(* IEC 61131-3 sources: plcassist-cli/packages/volt-lsp-iec/test-corpus/bakon-nano/Device/Plc Logic/Application/Library Manager/L_TF2P_TechModulesFollowingPositioning, 28 files *)

(* ---- L_TF2P_CONSTANTS.gvl ---- *)
VAR_GLOBAL
	GC_DWCHECKIDTAPPETREF : DWORD := 16#DC34;
	GC_LREPSILON : LREAL := 1E-06;
	GC_POSITIVE_LIMIT_32BIT : LREAL := 2147483647;
	GC_NEGATIVE_LIMIT_32BIT : LREAL := -2147483647;
	GC_PI : LREAL := 3.1415926535897931;
END_VAR

(* ---- L_TF2P_IACCESSPOINTS.itf ---- *)
INTERFACE L_TF2P_IACCESSPOINTS
END_INTERFACE

METHOD GET_PAP : POINTER TO L_TF2P_scAP_TM_TablePositioningBase
END_METHOD

(* ---- L_TF2P_ICONNECTORTABLEPOS.itf ---- *)
INTERFACE L_TF2P_ICONNECTORTABLEPOS
END_INTERFACE

(* ---- L_TF2P_ITABLEPOSITIONINGBASE.itf ---- *)
INTERFACE L_TF2P_ITABLEPOSITIONINGBASE
END_INTERFACE

METHOD PROFILEGENERATOR
VAR_INPUT
	ITFTECHMODULE : L_TF2P_ITablePositioningBase;
	XEXECUTE : BOOL;
	XCONTINUOUSUPDATE : BOOL;
	LRPOSITION : LREAL;
	LRVELOCITY : LREAL;
	LRENDVELOCITY : LREAL;
	LRACCELERATION : LREAL;
	LRDECELERATION : LREAL;
	LRJERK : LREAL;
	XPOSMODE : BOOL;
	EDIRECTION : MC_DIRECTION;
	EFUNCTIONTYP : L_MC1P_TypeFunction;
END_VAR
VAR_OUTPUT
	XDONE : BOOL;
	XBUSY : BOOL;
	XACTIVE : BOOL;
	XCOMMANDABORTED : BOOL;
	XERROR : BOOL;
	EERRORID : L_IE1P_Error;
END_VAR
VAR_IN_OUT
	AXIS : AXIS_REF;
END_VAR
END_METHOD

(* ---- GETBOOLEANPROPERTY.fun ---- *)
FUNCTION GETBOOLEANPROPERTY : BOOL
VAR_INPUT
	STKEY : WSTRING;
END_VAR
END_FUNCTION

(* ---- GETCOMPANY.fun ---- *)
FUNCTION GETCOMPANY : WSTRING
END_FUNCTION

(* ---- GETNUMBERPROPERTY.fun ---- *)
FUNCTION GETNUMBERPROPERTY : DINT
VAR_INPUT
	STKEY : WSTRING;
END_VAR
END_FUNCTION

(* ---- GETTEXTPROPERTY.fun ---- *)
FUNCTION GETTEXTPROPERTY : WSTRING
VAR_INPUT
	STKEY : WSTRING;
END_VAR
END_FUNCTION

(* ---- GETTEXTPROPERTY2.fun ---- *)
FUNCTION GETTEXTPROPERTY2 : POINTER TO WSTRING
VAR_INPUT
	STKEY : WSTRING;
END_VAR
END_FUNCTION

(* ---- GETTITLE.fun ---- *)
FUNCTION GETTITLE : WSTRING
END_FUNCTION

(* ---- GETVERSION.fun ---- *)
FUNCTION GETVERSION : VERSION
END_FUNCTION

(* ---- GETVERSIONPROPERTY.fun ---- *)
FUNCTION GETVERSIONPROPERTY : VERSION
VAR_INPUT
	STKEY : WSTRING;
END_VAR
END_FUNCTION

(* ---- L_TF2P_CHECKEXTERNALBYLIMITER.fun ---- *)
FUNCTION L_TF2P_CHECKEXTERNALBYLIMITER : BOOL
VAR_INPUT
	DWLIMITERCONTROL : DWORD;
END_VAR
VAR_IN_OUT
	AXIS : AXIS_REF;
END_VAR
END_FUNCTION

(* ---- L_TF2P_GETSTARTMOVETOTARGETPOS.fun ---- *)
FUNCTION L_TF2P_GETSTARTMOVETOTARGETPOS : BOOL
VAR_INPUT
	MASTERVALUES : L_MC1P_IAXIS_REF_MASTERVALUES;
	LRSYNCDEC : LREAL;
	LRSYNCJERK : LREAL;
	LRTARGETPOS : LREAL;
END_VAR
VAR_IN_OUT
	AXIS : AXIS_REF;
END_VAR
END_FUNCTION

(* ---- L_TF2P_POSITIONINSIDEWINDOW.fun ---- *)
FUNCTION L_TF2P_POSITIONINSIDEWINDOW : BOOL
VAR_INPUT
	LRPOSIN : LREAL;
	LRLOWERWINDOW : LREAL;
	LRUPPERWINDOW : LREAL;
END_VAR
VAR_OUTPUT
	XERROR : BOOL := FALSE;
END_VAR
VAR_IN_OUT
	AXIS : AXIS_REF;
END_VAR
END_FUNCTION

(* ---- GLOBALTEXTLIST.fb ---- *)
FUNCTION_BLOCK GLOBALTEXTLIST
VAR
	M_TEXTLISTFILE : STRING(255);
	_STNAMESPACE : STRING;
END_VAR
END_FUNCTION_BLOCK

(* ---- L_TB2A_PROFILEMANAGER.fb ---- *)
FUNCTION_BLOCK L_TB2A_PROFILEMANAGER
VAR_INPUT
	XEXECUTE : BOOL;
	XABORT : BOOL;
	WSTARTNUMBER : WORD;
	XNEXTPROFILE : BOOL;
END_VAR
VAR_OUTPUT
	XBUSY : BOOL;
	XDONE : BOOL;
	XABORTED : BOOL;
	XERROR : BOOL;
	EERRORID : L_IE1P_Error;
	XPROFILEERROR : BOOL;
	EPROFILEERRORID : L_IE1P_Error;
	WACTPROFILE : WORD;
	PACTPROFILE : POINTER TO L_TF2P_scPositionProfile;
	XHASNEXT : BOOL;
	XRTRIG : BOOL;
	EPROFILETYPE : L_MC1P_TypeFunction;
	XMOVEABS : BOOL;
	XMOVEREL : BOOL;
	XMOVEVEL : BOOL;
	XMOVECONTABS : BOOL;
	XMOVECONTREL : BOOL;
	XTPINSIDEWINDOW : BOOL;
	XTPOUTSIDEWINDOW : BOOL;
	XTPMISSED : BOOL;
	EDIRECTION : MC_DIRECTION;
END_VAR
VAR_IN_OUT
	ASCPROFILES : ARRAY [1..15] OF L_TF2P_scPositionProfile;
	SCTPRECDATA : L_MC1P_TpReceiveData;
	AXIS : AXIS_REF;
END_VAR
VAR
	_MODEL : L_UBUP_BehaviourModel_ETrigA;
	_XNEXTPROFILETRIG : R_TRIG;
	_XTPPROFILE : R_TRIG;
	LRTP_RELDIFF : LREAL;
	XTPWINDOWOPENED : BOOL;
	XTPWINDOWOPEN : BOOL;
	XTP_REL_PROFILEACTIVE : BOOL;
END_VAR
END_FUNCTION_BLOCK

METHOD CYCLICACTION
VAR_INPUT
	ITFTIMINGCONTROLLER : L_UBUP_ITimingController;
END_VAR
VAR_OUTPUT
	XCOMPLETE : BOOL;
	XABORT : BOOL;
	IERRORID : INT;
END_VAR
END_METHOD

METHOD FINALIZEACTION
VAR_INPUT
	XABORTPROPOSED : BOOL;
	IERRORIDPROPOSED : INT;
END_VAR
VAR_OUTPUT
	XCOMPLETE : BOOL;
	XABORT : BOOL;
	IERRORID : INT;
END_VAR
END_METHOD

METHOD RESETACTION
VAR_OUTPUT
	XCOMPLETE : BOOL;
END_VAR
END_METHOD

METHOD STARTACTION
VAR_OUTPUT
	XCOMPLETE : BOOL;
	IERRORID : INT;
END_VAR
END_METHOD

METHOD FB_INIT : BOOL
VAR_INPUT
	BINITRETAINS : BOOL;
	BINCOPYCODE : BOOL;
END_VAR
END_METHOD

METHOD GET_POSITIONINGMODE
VAR_OUTPUT
	EERRORID : L_IE1P_Error;
END_VAR
END_METHOD

METHOD GET_PROFILE
END_METHOD

METHOD GET_TPDETECTION
VAR_OUTPUT
	EERRORID : L_IE1P_Error;
END_VAR
END_METHOD

(* ---- L_TF2P_CONDITIONPROFILEMANAGER.fb ---- *)
FUNCTION_BLOCK L_TF2P_CONDITIONPROFILEMANAGER EXTENDS L_UBUP_ConditionBase
VAR_INPUT
	EPOSITIONINGMODE : L_TF2P_ePositioningMode;
	EINVALIDPROFILEID : L_IE1P_Error;
	EACTSTATE : L_TB2P_States;
END_VAR
VAR_IN_OUT
	AXIS : AXIS_REF;
END_VAR
END_FUNCTION_BLOCK

METHOD VERIFY : BOOL
VAR_OUTPUT
	XCONDITIONERROR : BOOL;
	EERRORIDPROPOSED : L_IE1P.L_IE1P_Error;
END_VAR
END_METHOD

(* ---- L_TF2P_CONTROLUNIT_ACTUALSPEED.fb ---- *)
FUNCTION_BLOCK L_TF2P_CONTROLUNIT_ACTUALSPEED
VAR_INPUT
	XENABLE : BOOL := FALSE;
	XENABLEOPERATION : BOOL := FALSE;
	XSPEEDCONTROL : BOOL := FALSE;
	SCPROFILELIMITS : L_TF2P_scProfileLimits;
	XENABLEEXTVEL : BOOL := FALSE;
	LREXTVEL : LREAL := 0;
	XENABLEEXTACCDECJERK : BOOL := FALSE;
	LREXTACC : LREAL := 0;
	LREXTDEC : LREAL := 0;
	LREXTJERK : LREAL := 0;
	XENABLEEXTTRQ : BOOL := FALSE;
	LREXTTRQ : LREAL := 0;
	XFASTSLOW : BOOL;
	XINVERTDIRECTION : BOOL;
	SCPROFILEACTUALSPEED : L_TF2P_scProfileDataState_int;
	XBRAKEISUSED : BOOL := FALSE;
	XBRAKERELEASED : BOOL := FALSE;
	ETMSTATES : L_TB2P_States;
	XAXISWARNING : BOOL;
	XTMERROR : BOOL;
	XSTO : BOOL;
	XAXISENABLED : BOOL := FALSE;
	XAXISREADY : BOOL := FALSE;
END_VAR
VAR_OUTPUT
	XENABLED : BOOL := FALSE;
	XBUSY : BOOL := FALSE;
	SCCONTROLUNIT : L_TF2P_scControlUnit;
	XERROR : BOOL;
	EERRORID : L_IE1P_Error;
	XEXTVELACTIVE : BOOL;
	XEXTTRQACTIVE : BOOL;
	XEXTACCDECJERKACTIVE : BOOL := FALSE;
	XMOVEVELEXECUTE : BOOL;
	XABORTOUT : BOOL;
	ESETDIRECTION : L_MC1P.MC_DIRECTION;
END_VAR
VAR_IN_OUT
	XNEWCOMMAND : BOOL;
END_VAR
VAR
	XNOTFIRSTCYCLE : BOOL := FALSE;
	XSPEEDCONTROL_OLD : BOOL;
END_VAR
END_FUNCTION_BLOCK

(* ---- L_TF2P_FOLLOWSETVALUESBASE.fb ---- *)
FUNCTION_BLOCK L_TF2P_FOLLOWSETVALUESBASE EXTENDS L_TB2P_TechModuleBase
VAR_INPUT
	XENABLE : BOOL;
	XENABLEOPERATION : BOOL;
	XRESETERROR : BOOL;
	XQSPAPPLICATION : BOOL;
	XABORT : BOOL;
	XJOGPOS : BOOL;
	XJOGNEG : BOOL;
	XHOMEEXECUTE : BOOL;
	LROVERRIDE : LREAL := 1;
	SCCTRLBASICMOTION : L_TB2P_scCtrlBasicMotion;
	SCPAR : L_TF2P_scPar_FollowSetValuesBase;
	SCACCESSPOINTS : L_TF2P_scAP_FollowSetValuesBase;
	XFOLLOWSETVALUES : BOOL;
	LRSETVELOCITY : LREAL;
	LRSETTORQUE : LREAL;
END_VAR
VAR_OUTPUT
	XREADYFOROPERATION : BOOL;
	XOPERATIONENABLED : BOOL;
	XREADYFORMOTION : BOOL;
	XERROR : BOOL;
	XWARNING : BOOL;
	EERRORID : L_IE1P_Error;
	XSTOACTIVE : BOOL;
	XQSPACTIVE : BOOL;
	XABORTBUSY : BOOL;
	XABORTDONE : BOOL;
	XJOGGINGBUSY : BOOL;
	XHOMINGBUSY : BOOL;
	XHOMINGDONE : BOOL;
	XISHOMED : BOOL;
	ETMSTATE : L_TB2P_States := L_TB2P_States.DISABLED;
	SCSTATUSBASICMOTION : L_TB2P_scStatusBasicMotion;
	LRACTVEL : LREAL;
	LRSETVELOUT : LREAL;
	LRACTPOS : LREAL;
	LRSETPOSOUT : LREAL;
	LRACTFOLLOWINGERROR : LREAL;
	SCSIGNALFLOW : L_TF2P_scSF_FollowSetValuesBase;
	XFOLLOWVELOCITYBUSY : BOOL;
	XFOLLOWTORQUEBUSY : BOOL;
	XVELLIMITACTIVE : BOOL;
	XACCDECLIMITACTIVE : BOOL;
	XTORQUEINTARGET : BOOL;
	LRACTTORQUE : LREAL;
	LRSETTORQUEOUT : LREAL;
END_VAR
VAR_IN_OUT
	AXIS : AXIS_REF;
END_VAR
VAR
	TM_INT : L_TF2P_TM_FollowSetValuesBase := STRUCT(ModuleHandler := ModuleHandler);
	XENABLE_OLD : BOOL;
	_UICALLMFUNIDXINPUT : UINT := 1;
	_UICALLMFUNIDXOUTPUT : UINT := 1;
	_ASCINPUT : ARRAY [1.._MCCall.c_BufferDepthInput] OF L_TF2P_FollowSetValuesBaseIn;
	_ASCOUTPUT : ARRAY [1.._MCCall.c_BufferDepthOutput] OF L_TF2P_FollowSetValuesBaseOut;
	_ASCPARCORE : ARRAY [1.._MCCall.c_BufferDepthInput] OF L_TF2P_scPar_FollowSetValuesBase;
	_ASCACCESSPOINTSCORE : ARRAY [1.._MCCall.c_BufferDepthInput] OF L_TF2P_scAP_FollowSetValuesBase;
	_ASCSIGNALFLOWCORE : ARRAY [1.._MCCall.c_BufferDepthOutput] OF L_TF2P_scSF_FollowSetValuesBase;
	_MCCALL : L_UM1P_MCCall;
	SCPAR_INT : L_TF2P_scPar_FollowSetValuesBase;
	_SCINPUTVISU : L_TF2P_FollowSetValuesBaseIn;
	_PSCINPUTVISU : POINTER TO L_TF2P_FollowSetValuesBaseIn := ADR(_scInputVisu);
	_PSCOUTPUTVISU : POINTER TO L_TF2P_FollowSetValuesBaseOut := ADR(_ascOutput[1]);
	_PSCPARVISU : POINTER TO L_TF2P_scPar_FollowSetValuesBase := ADR(scPar_int);
	ITFITECHMODULEINTERNAL : L_TB2P_ITechModuleInternal;
	LRJERKDEC : LREAL;
	LRJOGGINGJERKDEC : LREAL;
	REMAININGTIMEOFPROFILE : LREAL;
	REMAININGTIMEOFPROFILEAVAILABLE : BOOL;
END_VAR
END_FUNCTION_BLOCK

METHOD GET_PAP : POINTER TO L_TB2P_scAP_TM_MotionControl
END_METHOD

METHOD GET_PPAR : POINTER TO L_TB2P.L_TB2P_scPar_TM_MotionControl
END_METHOD

METHOD GET_PSF : POINTER TO L_TB2P_scSF_TM_MotionControl
END_METHOD

METHOD CALLFUNCTION
VAR_INPUT
	UIINPUTDATAIDX : UINT;
	UIOUTPUTDATAIDX : UINT;
END_VAR
END_METHOD

METHOD COPYINPUTS : BOOL
VAR_INPUT
	IDX : WORD;
END_VAR
END_METHOD

METHOD COPYOUTPUTS : BOOL
VAR_INPUT
	IDX : WORD;
END_VAR
END_METHOD

METHOD FUNCTIONWASCALLEDTWICE : BOOL
VAR_INPUT
	IDX : WORD;
END_VAR
END_METHOD

METHOD HANDLESTANDARDCALL : BOOL
END_METHOD

METHOD SYNCOUTPUTS
VAR_INPUT
	UICOPYOUTPUTFROMIDX : UINT;
	UICOPYOUTPUTTOIDX : UINT;
END_VAR
END_METHOD

METHOD CALL_INTERNALCTRL
END_METHOD

(* ---- L_TF2P_SPEEDCONTROLBASE.fb ---- *)
FUNCTION_BLOCK L_TF2P_SPEEDCONTROLBASE EXTENDS L_TB2P_TechModuleBase
VAR_INPUT
	XENABLE : BOOL;
	XENABLEOPERATION : BOOL;
	XRESETERROR : BOOL;
	XQSPAPPLICATION : BOOL;
	XABORT : BOOL;
	XJOGPOS : BOOL;
	XJOGNEG : BOOL;
	XHOMEEXECUTE : BOOL;
	LROVERRIDE : LREAL := 1;
	SCCTRLBASICMOTION : L_TB2P_scCtrlBasicMotion;
	SCPAR : L_TF2P_scPar_SpeedControlBase;
	SCACCESSPOINTS : L_TF2P_scAP_SpeedControlBase;
	XSPEEDCONTROL : BOOL;
	XNEGATIVEDIRECTION : BOOL;
	LRSETVEL : LREAL;
	XUSEEXTACCDECJERK : BOOL;
	LREXTACC : LREAL := 100;
	LREXTDEC : LREAL := 100;
	LREXTJERK : LREAL := 100000;
	LRSETOFFSETVEL : LREAL := 0.0;
	XUSEPROFILEVEL : BOOL;
	WPROFILENUMBER : WORD;
END_VAR
VAR_OUTPUT
	XREADYFOROPERATION : BOOL;
	XOPERATIONENABLED : BOOL;
	XREADYFORMOTION : BOOL;
	XERROR : BOOL;
	XWARNING : BOOL;
	EERRORID : L_IE1P_Error;
	XSTOACTIVE : BOOL;
	XQSPACTIVE : BOOL;
	XABORTBUSY : BOOL;
	XABORTDONE : BOOL;
	XJOGGINGBUSY : BOOL;
	XHOMINGBUSY : BOOL;
	XHOMINGDONE : BOOL;
	XISHOMED : BOOL;
	ETMSTATE : L_TB2P_States := L_TB2P_States.DISABLED;
	SCSTATUSBASICMOTION : L_TB2P_scStatusBasicMotion;
	LRACTVEL : LREAL;
	LRSETVELOUT : LREAL;
	LRACTPOS : LREAL;
	LRSETPOSOUT : LREAL;
	LRACTFOLLOWINGERROR : LREAL;
	SCSIGNALFLOW : L_TF2P_scSF_SpeedControlBase;
	XSPEEDCONTROLBUSY : BOOL;
	XEXTACCDECJERKACTIVE : BOOL;
	XOFFSETVELACTIVE : BOOL;
	XPROFILEVELACTIVE : BOOL;
	WACTIVEPROFILE : WORD;
END_VAR
VAR_IN_OUT
	AXIS : AXIS_REF;
END_VAR
VAR
	TM_INT : L_TF2P_TM_SpeedControlBase := STRUCT(ModuleHandler := ModuleHandler);
	PPAR : POINTER TO L_TF2P_scPar_SpeedControlBase;
	PPAR_INT : POINTER TO L_TF2P_scPar_SpeedControlBase;
	_UICALLMFUNIDXINPUT : UINT := 1;
	_UICALLMFUNIDXOUTPUT : UINT := 1;
	_ASCINPUT : ARRAY [1.._MCCall.c_BufferDepthInput] OF L_TF2P_SpeedControlBaseIn;
	_ASCOUTPUT : ARRAY [1.._MCCall.c_BufferDepthOutput] OF L_TF2P_SpeedControlBaseOut;
	_ASCPARCORE : ARRAY [1.._MCCall.c_BufferDepthInput] OF L_TF2P_scPar_SpeedControlBase;
	_ASCACCESSPOINTSCORE : ARRAY [1.._MCCall.c_BufferDepthInput] OF L_TF2P_scAP_SpeedControlBase;
	_ASCSIGNALFLOWCORE : ARRAY [1.._MCCall.c_BufferDepthOutput] OF L_TF2P_scSF_SpeedControlBase;
	_MCCALL : L_UM1P_MCCall;
	SCPAR_INT : L_TF2P_scPar_SpeedControlBase;
	_SCINPUTVISU : L_TF2P_SpeedControlBaseIn;
	_PSCINPUTVISU : POINTER TO L_TF2P_SpeedControlBaseIn := ADR(_scInputVisu);
	_PSCOUTPUTVISU : POINTER TO L_TF2P_SpeedControlBaseOut := ADR(_ascOutput[1]);
	_PSCPARVISU : POINTER TO L_TF2P_scPar_SpeedControlBase := ADR(scPar_int);
	XVISPOINTMIN : BOOL;
	XVISPOINTMAX : BOOL;
	XVISUSETPOSUP : BOOL;
	XVISUSETPOSDOWN : BOOL;
	RTRIGUP : R_TRIG;
	RTRIGDOWN : R_TRIG;
	IMAXPOINTS : INT := 11;
	IPOINT : INT := 0;
	ITFITECHMODULEINTERNAL : L_TB2P_ITechModuleInternal;
	LRJERKDEC : LREAL;
	LRJOGGINGJERKDEC : LREAL;
	REMAININGTIMEOFPROFILE : LREAL;
	REMAININGTIMEOFPROFILEAVAILABLE : BOOL;
END_VAR
END_FUNCTION_BLOCK

METHOD GET_PAP : POINTER TO L_TB2P_scAP_TM_MotionControl
END_METHOD

METHOD GET_PPAR : POINTER TO L_TB2P.L_TB2P_scPar_TM_MotionControl
END_METHOD

METHOD GET_PSF : POINTER TO L_TB2P_scSF_TM_MotionControl
END_METHOD

METHOD CALLFUNCTION
VAR_INPUT
	UIINPUTDATAIDX : UINT;
	UIOUTPUTDATAIDX : UINT;
END_VAR
END_METHOD

METHOD COPYINPUTS : BOOL
VAR_INPUT
	IDX : WORD;
END_VAR
END_METHOD

METHOD COPYOUTPUTS : BOOL
VAR_INPUT
	IDX : WORD;
END_VAR
END_METHOD

METHOD FUNCTIONWASCALLEDTWICE : BOOL
VAR_INPUT
	IDX : WORD;
END_VAR
END_METHOD

METHOD HANDLESTANDARDCALL : BOOL
END_METHOD

METHOD SYNCOUTPUTS
VAR_INPUT
	UICOPYOUTPUTFROMIDX : UINT;
	UICOPYOUTPUTTOIDX : UINT;
END_VAR
END_METHOD

METHOD CALL_INTERNALCTRL
END_METHOD

METHOD CALL_VISUPROFILES
END_METHOD

(* ---- L_TF2P_TABLEPOSITIONINGBASE.fb ---- *)
FUNCTION_BLOCK L_TF2P_TABLEPOSITIONINGBASE EXTENDS L_TB2P_TechModuleBase
VAR_INPUT
	XUSEORIGINAL : BOOL;
	XENABLE : BOOL;
	XENABLEOPERATION : BOOL;
	XRESETERROR : BOOL;
	XQSPAPPLICATION : BOOL;
	XABORT : BOOL;
	XJOGPOS : BOOL;
	XJOGNEG : BOOL;
	XHOMEEXECUTE : BOOL;
	LROVERRIDE : LREAL := 1;
	SCCTRLBASICMOTION : L_TB2P_scCtrlBasicMotion;
	SCPAR : L_TF2P_scPar_TablePositioningBase;
	SCACCESSPOINTS : L_TF2P_scAP_TablePositioningBase;
	WPROFILENUMBER : WORD := 1;
	XEXECUTEPOSITIONING : BOOL;
	SCTPRECDATA : L_MC1P_TpReceiveData;
END_VAR
VAR_OUTPUT
	XREADYFOROPERATION : BOOL;
	XOPERATIONENABLED : BOOL;
	XREADYFORMOTION : BOOL;
	XERROR : BOOL;
	XWARNING : BOOL;
	EERRORID : L_IE1P_Error;
	XSTOACTIVE : BOOL;
	XQSPACTIVE : BOOL;
	XABORTBUSY : BOOL;
	XABORTDONE : BOOL;
	XJOGGINGBUSY : BOOL;
	XHOMINGBUSY : BOOL;
	XHOMINGDONE : BOOL;
	XISHOMED : BOOL;
	ETMSTATE : L_TB2P_States;
	SCSTATUSBASICMOTION : L_TB2P_scStatusBasicMotion;
	LRACTVEL : LREAL;
	LRSETVELOUT : LREAL;
	LRACTPOS : LREAL;
	LRSETPOSOUT : LREAL;
	LRACTFOLLOWINGERROR : LREAL;
	SCSIGNALFLOW : L_TF2P_scSF_TablePositioningBase;
	XPROFILEBUSY : BOOL;
	XPROFILEDONE : BOOL;
	XDRIVEINTARGET : BOOL;
	WACTIVEPROFILE : WORD;
END_VAR
VAR_IN_OUT
	AXIS : AXIS_REF;
END_VAR
VAR
	XUSEORIGINAL_OLD : BOOL;
	ITFCONNECTORTABLEPOS : L_TF2P_IConnectorTablePos;
	TM_INT : L_TF2P_TM_TablePositioningBase;
	SCPAR_INT : L_TF2P_scPar_TablePositioningBase;
	SCSIGNALFLOW_INT : L_TF2P_scSF_TablePositioningBase;
	IPOINT : INT := 1;
	_UICALLMFUNIDXINPUT : UINT := 1;
	_UICALLMFUNIDXOUTPUT : UINT := 1;
	_MCCALL : L_UM1P_MCCall;
	_ASCINPUT : ARRAY [1.._MCCall.c_BufferDepthInput] OF L_TF2P_TablePositioningBaseIn;
	_ASCOUTPUT : ARRAY [1.._MCCall.c_BufferDepthOutput] OF L_TF2P_TablePositioningBaseOut;
	_ASCPARCORE : ARRAY [1.._MCCall.c_BufferDepthInput] OF L_TF2P_scPar_TablePositioningBase;
	_ASCACCESSPOINTSCORE : ARRAY [1.._MCCall.c_BufferDepthInput] OF L_TF2P_scAP_TablePositioningBase;
	_ASCSIGNALFLOWCORE : ARRAY [1.._MCCall.c_BufferDepthOutput] OF L_TF2P_scSF_TablePositioningBase;
	_SCINPUTVISU : L_TF2P_TablePositioningBaseIn;
	_PSCINPUTVISU : POINTER TO L_TF2P_TablePositioningBaseIn := ADR(_scInputVisu);
	_PSCOUTPUTVISU : POINTER TO L_TF2P_TablePositioningBaseOut := ADR(_ascOutput[1]);
	_PSCPARVISU : POINTER TO L_TF2P_scPar_TablePositioningBase := ADR(scPar_int);
	ITFBASICMOTIONBASE : L_TB2P.L_TB2P_IBasicMotionBase;
	ITFITECHMODULEINTERNAL : L_TB2P_ITechModuleInternal;
	ITFTABLEPOSITIONING : L_TF2P_ITablePositioningBase;
	LRJERKDEC : LREAL;
	LRJOGGINGJERKDEC : LREAL;
	REMAININGTIMEOFPROFILE : LREAL;
	REMAININGTIMEOFPROFILEAVAILABLE : BOOL;
END_VAR
END_FUNCTION_BLOCK

METHOD CALL_ABC
VAR_INPUT
	ITFTECHMODULE : L_TB2P.L_TB2P_IBasicMotionBase;
	XQSPAPPLICATION : BOOL;
	XHALT : BOOL;
	XABORT : BOOL;
	XHOMEEXECUTE : BOOL;
	XJOGPOS : BOOL;
	XJOGNEG : BOOL;
	XFINISHPOSITIONING : BOOL;
	XMOVEVELEXECUTE : BOOL;
	XMOVEABSEXECUTE : BOOL;
	XMOVERELEXECUTE : BOOL;
	XENABLEOPERATION : BOOL;
	XRESETERROR : BOOL;
	XENABLEPOSITIVE : BOOL;
	XENABLENEGATIVE : BOOL;
	XDISABLESWLIMIT : BOOL;
	LROVERRIDE : LREAL;
	LROVERRIDEACC : LREAL;
	LROVERRIDEJERK : LREAL;
	XRESETHOMEPOSITION : BOOL;
	XCONTINUOUSUPDATE : BOOL;
	LRPOS_DIST : LREAL;
	LRVEL : LREAL;
	LRACC : LREAL;
	LRDEC : LREAL;
	LRJERK : LREAL;
	EDIRECTION : L_TB2P.MC_DIRECTION;
	SCHOMEEXTTP : L_TB2P.MC_TRIGGER_REF;
	XHOMEABSSWITCH : BOOL;
	XSPECIALABORTBEHAVIOR : BOOL;
	LRABORTDEC : LREAL;
	LRABORTJERK : LREAL;
END_VAR
VAR_OUTPUT
	XERROR : BOOL;
	EERRORID : L_TB2P.L_IE1P_Error;
	XFUNBUSY : BOOL;
	XFUNDONE : BOOL;
	XFUNCOMMANDABORTED : BOOL;
	EFUNSTATEACT : L_TB2P.L_MC1P_ABC_State;
	ECONTROLMODE : L_TB2P.L_MC1P_ControlMode;
	XISHOMED : BOOL;
	XHWLIMITSWITCHNEG : BOOL;
	XHWLIMITSWITCHPOS : BOOL;
	XSWLIMITENABLED : BOOL;
	XSWLIMITSWITCHNEG : BOOL;
	XSWLIMITSWITCHPOS : BOOL;
	EAXISTYPE : L_TB2P.L_MC1P_DriveType;
	EAXISSTATE : L_TB2P.L_MC1P_AXIS_STATE;
	XSTOACTIVE : BOOL;
	XREADYFOROPERATION : BOOL;
	XOPERATIONENABLED : BOOL;
	XREADYFORMOTION : BOOL;
	XAXISWARNING : BOOL;
	XAXISERROR : BOOL;
	EAXISERRORID : L_TB2P.L_IE1P_Error;
	XDRIVEWARNING : BOOL;
	XDRIVEERROR : BOOL;
	DWDRIVEERRORID : DWORD;
	LRACTPOS : LREAL;
	LRACTVEL : LREAL;
	LRSETPOSOUT : LREAL;
	LRSETVELOUT : LREAL;
	LRACTFOLLOWINGERROR : LREAL;
	XINPOSITION : BOOL;
	XSTANDSTILLSETVELOCITY : BOOL;
	XSTANDSTILLACTVELOCITY : BOOL;
	XCONSTANTVELOCITY : BOOL;
	XACCELERATING : BOOL;
	XDECELERATING : BOOL;
	XDIRECTIONPOSITIVE : BOOL;
	XDIRECTIONNEGATIVE : BOOL;
	XAXISAVAILABLE : BOOL;
END_VAR
VAR_IN_OUT
	AXIS : AXIS_REF;
END_VAR
END_METHOD

METHOD GET_PAP : POINTER TO L_TB2P_scAP_TM_MotionControl
END_METHOD

METHOD GET_PPAR : POINTER TO L_TB2P.L_TB2P_scPar_TM_MotionControl
END_METHOD

METHOD GET_PSF : POINTER TO L_TB2P_scSF_TM_MotionControl
END_METHOD

METHOD PROFILEGENERATOR
VAR_INPUT
	ITFTECHMODULE : L_TF2P_ITablePositioningBase;
	XEXECUTE : BOOL;
	XCONTINUOUSUPDATE : BOOL;
	LRPOSITION : LREAL;
	LRVELOCITY : LREAL;
	LRENDVELOCITY : LREAL;
	LRACCELERATION : LREAL;
	LRDECELERATION : LREAL;
	LRJERK : LREAL;
	XPOSMODE : BOOL;
	EDIRECTION : MC_DIRECTION;
	EFUNCTIONTYP : L_MC1P_TypeFunction;
END_VAR
VAR_OUTPUT
	XDONE : BOOL;
	XBUSY : BOOL;
	XACTIVE : BOOL;
	XCOMMANDABORTED : BOOL;
	XERROR : BOOL;
	EERRORID : L_IE1P_Error;
END_VAR
VAR_IN_OUT
	AXIS : AXIS_REF;
END_VAR
END_METHOD

METHOD CALLFUNCTION
VAR_INPUT
	UIINPUTDATAIDX : UINT;
	UIOUTPUTDATAIDX : UINT;
END_VAR
END_METHOD

METHOD COPYINPUTS : BOOL
VAR_INPUT
	IDX : WORD;
END_VAR
END_METHOD

METHOD COPYOUTPUTS : BOOL
VAR_INPUT
	IDX : WORD;
END_VAR
END_METHOD

METHOD FUNCTIONWASCALLEDTWICE : BOOL
VAR_INPUT
	IDX : WORD;
END_VAR
END_METHOD

METHOD HANDLESTANDARDCALL : BOOL
END_METHOD

METHOD SYNCOUTPUTS
VAR_INPUT
	UICOPYOUTPUTFROMIDX : UINT;
	UICOPYOUTPUTTOIDX : UINT;
END_VAR
END_METHOD

METHOD FB_INIT : BOOL
VAR_INPUT
	BINITRETAINS : BOOL;
	BINCOPYCODE : BOOL;
END_VAR
END_METHOD

METHOD CALL_INTERNALCTRL
END_METHOD

(* ---- L_TF2P_TM_FOLLOWSETVALUESBASE.fb ---- *)
FUNCTION_BLOCK L_TF2P_TM_FOLLOWSETVALUESBASE EXTENDS L_TB2P_TM_MotionControl
VAR
	TM_FOLLOWSETVALUESBASECONFIG : L_TB2P_ModuleHandlerConfig;
	PSCINPUT : POINTER TO L_TF2P_FollowSetValuesBaseIn;
	PSCOUTPUT : POINTER TO L_TF2P_FollowSetValuesBaseOut;
	PPAR : POINTER TO L_TF2P_scPar_TM_FollowSetValuesBase;
	PSF : POINTER TO L_TF2P_scSF_TM_FollowSetValuesBase;
	PAP : POINTER TO L_TF2P_scAP_TM_FollowSetValuesBase;
	SCPAR_INT : L_TF2P_scPar_TM_FollowSetValuesBase;
	LRFILTERTIMEFACTOR : LREAL;
	LRSETVALUEFILTERED : LREAL;
	LRRAMPGEN_SETVALUEOUT : LREAL;
	LRTASKCYCLE : LREAL;
	LRFILTERTIME : LREAL;
	LRTIME : LREAL;
	LRSETVALUE : LREAL;
	WLENZESTATUSWORD : WORD;
	XVELLIMITSERR : BOOL;
	XVELLIMITSWRN : BOOL;
	IACTMASTERDIRECTION_INT : INT;
	XTM_ABORT : BOOL;
	XTM_ABORTNEXTCYCLE : BOOL;
	XWARNINGDIRECTIONDISABLED : BOOL;
	FB_READHALTDEC : MC_ReadParameter := STRUCT(ParameterNumber := 186);
	FB_READHALTJERK : MC_ReadParameter := STRUCT(ParameterNumber := 187);
	LRHALTDEC_INT : LREAL;
	LRHALTJERK_INT : LREAL;
	L_MC1P_FOLLOWSETVALUES1 : L_MC1P_FollowSetValues := STRUCT(UseSpeedCtrlMode := TRUE);
	L_MC1P_TORQUECONTROL1 : L_MC1P_TorqueControl;
	L_MC1P_RAMPGENERATOR1 : L_MC1P_RampGenerator;
END_VAR
END_FUNCTION_BLOCK

METHOD CALL_ALLOCPOINTADR
END_METHOD

METHOD CALL_ERRORRESETACTIVE
END_METHOD

METHOD CALL_ERRORHANDLER
END_METHOD

METHOD CALL_FBMETHODS
END_METHOD

METHOD CALL_FB_READHALTDEC
END_METHOD

METHOD CALL_FB_READHALTJERK
END_METHOD

METHOD CALL_INITDONE
END_METHOD

METHOD CALL_INITROUTINE
END_METHOD

METHOD CALL_INTERNALCTRL
END_METHOD

METHOD CALL_OUTPUT
END_METHOD

METHOD CALL_OUTPUT_SF
END_METHOD

METHOD CALL_PT1FILTER
END_METHOD

METHOD CALL_RAMPGENERATOR
END_METHOD

METHOD CALL_REQUESTS_EXT
END_METHOD

METHOD CALL_RESETCOMMANDS
END_METHOD

METHOD CALL_RESETOUTPUT
END_METHOD

METHOD CALL_SPEEDCONTROL
END_METHOD

METHOD CALL_TORQUECONTROL
END_METHOD

METHOD CALL_ABC
END_METHOD

METHOD CALL_ABC_INPUT
END_METHOD

METHOD CALL_ABC_INPUT_PROFILEPARAMETER
END_METHOD

METHOD CALL_S042_ABORT_VELOCITYFOLLOWING
END_METHOD

METHOD CALL_S042_VELOCITYFOLLOWING
END_METHOD

METHOD CALL_S043_TORQUEFOLLOWING
END_METHOD

METHOD CALL_STATEMACHINE
END_METHOD

METHOD CALL_T000_ALLSTATES
END_METHOD

METHOD MAPTMSTATE
VAR_INPUT
	ETMSTATEINTERNAL : L_TB2P_States;
END_VAR
VAR_OUTPUT
	ETMSTATEEXTERNAL : L_TB2P_States;
END_VAR
END_METHOD

METHOD CALL_T000_ALLSTATES_OUT
END_METHOD

(* ---- L_TF2P_TM_SPEEDCONTROLBASE.fb ---- *)
FUNCTION_BLOCK L_TF2P_TM_SPEEDCONTROLBASE EXTENDS L_TB2P_TM_MotionControl
VAR
	TM_SPEEDCONTROLBASE : L_TB2P_ModuleHandlerConfig;
	PSCINPUT : POINTER TO L_TF2P_SpeedControlBaseIn;
	PSCOUTPUT : POINTER TO L_TF2P_SpeedControlBaseOut;
	PPAR : POINTER TO L_TF2P_scPar_TM_SpeedControlBase;
	PSF : POINTER TO L_TF2P_scSF_TM_SpeedControlBase;
	PAP : POINTER TO L_TF2P_scAP_TM_SpeedControlBase;
	SCPAR_INT : L_TF2P_scPar_TM_SpeedControlBase;
	XSPEEDCONTROLACTIVE_INT : BOOL;
	XSPEEDCONTROLBUSY_INT : BOOL;
	XCOMMANDABORTED_INT : BOOL;
	XNEWCOMMAND : BOOL;
	XHALT_LINKED : BOOL;
	XCU_ABORT_OLD : BOOL;
	XABORT_INT_OLD : BOOL;
	XQSPAPPLICATION_INT_OLD : BOOL;
	XSPEEDCONTROL_INT_OLD : BOOL;
	XCU_MOVEVELEXECUTE_INT_OLD : BOOL;
	ECONTROLMODE_OLD : L_MC1P_ControlModeSet;
	XABC_MOVEVELEXECUTE_OLD : BOOL;
	FB_CU_ACTUALSPEED : L_TF2P_ControlUnit_ActualSpeed;
	FB_BRAKEINTERFACE : L_MC1P_BrakeInterface;
	FB_SR_XHALT : SR;
	XUSEPROFILEDATA : BOOL;
	XFUNDONESPEEDCONTROL : BOOL;
	XINVALIDPROFILE_INT : BOOL;
	XWARNINGINVALIDPROFILE_INT : BOOL;
	XERRORINVALIDPROFILE_INT : BOOL;
	WPROFILEINDEXMIN : WORD := 0;
	WPROFILEINDEXMAX : WORD := 15;
END_VAR
END_FUNCTION_BLOCK

METHOD CALL_ALLOCPOINTADR
END_METHOD

METHOD CALL_BRAKEINTERFACE
END_METHOD

METHOD CALL_CU_ACTUALSPEED
END_METHOD

METHOD CALL_CU_ACTUALSPEED_INPUT
END_METHOD

METHOD CALL_ERRORHANDLER
END_METHOD

METHOD CALL_INITDONE
END_METHOD

METHOD CALL_INITROUTINE
END_METHOD

METHOD CALL_INTERNALCTRL
END_METHOD

METHOD CALL_OUTPUT
END_METHOD

METHOD CALL_OUTPUT_SF
END_METHOD

METHOD CALL_REQUESTS_EXT
END_METHOD

METHOD CALL_RESETCOMMANDS
END_METHOD

METHOD CALL_RESETOUTPUT
END_METHOD

METHOD CALL_ABC_INPUT
END_METHOD

METHOD CALL_ABC_INPUT_PROFILEPARAMETER
END_METHOD

METHOD CALL_S002_STANDBY
END_METHOD

METHOD CALL_S010_JOGGING
END_METHOD

METHOD CALL_S013_MOVEVEL
END_METHOD

METHOD CALL_S017_EXTERNAL
END_METHOD

METHOD CALL_S999_ERROR
END_METHOD

METHOD CALL_STATEMACHINE
END_METHOD

METHOD CALL_T000_ALLSTATES
END_METHOD

METHOD CALL_S000_CYCLIC_OUT
END_METHOD

METHOD CALL_S014_MOVEABS_OUT
END_METHOD

METHOD CALL_S015_MOVEREL_OUT
END_METHOD

METHOD CALL_S017_EXTERNAL_OUT
END_METHOD

METHOD CALL_S996_STOP_OUT
END_METHOD

METHOD CALL_S999_ERROR_OUT
END_METHOD

(* ---- L_TF2P_TM_TABLEPOSITIONINGBASE.fb ---- *)
FUNCTION_BLOCK L_TF2P_TM_TABLEPOSITIONINGBASE EXTENDS L_TB2M_TM_MotionControl
VAR
	TM_TABLEPOS : L_TB2P_ModuleHandlerConfig;
	ITFPOSITIONINGBASE : L_TF2P_ITablePositioningBase := THIS^;
	SCDATA_INT : L_TF2P_scData_TM_TablePositioningBase;
	PDATA : POINTER TO L_TF2P_scData_TM_TablePositioningBase := ADR(scData_Int);
	PPAR : POINTER TO L_TF2P_scPar_TM_TablePositioningBase;
	PSF : POINTER TO L_TF2P_scSF_TM_TablePositioningBase;
	PAP : POINTER TO L_TF2P_scAP_TM_TablePositioningBase;
	PINPUT : POINTER TO L_TF2P_TablePositioningBaseIn;
	POUTPUT : POINTER TO L_TF2P_TablePositioningBaseOut;
	_SCTPRECDATA : L_MC1P_TpReceiveData;
	_FB_TPRECDATAPROXY : L_MC1P_TouchProbeRecDataProxy;
	FB_CONDITIONPROFILEMANAGER : L_TF2P_ConditionProfileManager;
	FB_CONDCOLLECTIONPROFILEMANAGER : L_UBUP_ConditionCollectionAND := STRUCT(aitfCondition := [fb_ConditionOperationEnabled, fb_ConditionProfileManager]);
	FB_CONDCOLLECTION : L_UBUP_ConditionCollectionAND := STRUCT(aitfCondition := [fb_ConditionOperationEnabled, fb_ConditionLimiter]);
	FB_CONDCOLLECTIONABSOLUTE : L_UBUP_ConditionCollectionAND := STRUCT(aitfCondition := [fb_CondCollection, fb_ConditionAxisHomed]);
	FB_TRANSITION2MOVEABSTABLEPOS : L_UBUP_RequestTransitionEdge;
	FB_TRANSITION2MOVEABSCONTTABLEPOS : L_UBUP_RequestTransitionEdge;
	FB_TRANSITION2MOVERELTABLEPOS : L_UBUP_RequestTransitionEdge;
	FB_TRANSITION2MOVERELCONTTABLEPOS : L_UBUP_RequestTransitionEdge;
	FB_TRANSITION2MOVEVELTABLEPOS : L_UBUP_RequestTransitionEdge;
	FB_TRANSITION2MOVEABSTABLEPOSFINISH : L_UBUP_RequestTransitionEdge;
	FB_TRANSITION2MOVEABSCONTTABLEPOSFINISH : L_UBUP_RequestTransitionEdge;
	FB_TRANSITION2MOVERELTABLEPOSFINISH : L_UBUP_RequestTransitionEdge;
	FB_TRANSITION2MOVERELCONTTABLEPOSFINISH : L_UBUP_RequestTransitionEdge;
	FB_TRANSITION2MOVEVELTABLEPOSFINISH : L_UBUP_RequestTransitionEdge;
	FB_TRANSITION2INVALIDPOSITIONINGMODE : L_UBUP_RequestTransitionLevel;
	FB_MOVEBASIC : L_MC1P_MoveBasic := STRUCT(wCalcProfileMode := 1);
	FB_PROFILEMANAGER : L_TB2A_ProfileManager;
	FB_DUMMYTEMPLATE : L_MC1P_Template_ForAxis;
	CONNECTOR : __SYSTEM.IQueryInterface;
	REMAININGTIMEOFPROFILE : LREAL;
	REMAININGTIMEOFPROFILEAVAILABLE : BOOL;
	TABLEPOSBASEEXTENSION : L_TF2P_ITablePositioningBase;
END_VAR
END_FUNCTION_BLOCK

METHOD CALLFBS
VAR_INPUT
	ECASE : L_UBUP_StateHandleCase;
END_VAR
END_METHOD

METHOD CALLSTATE
VAR_INPUT
	ITFSTATESERVER : L_UBUP_IStateServer;
	ISTATE : INT;
	ECASE : L_UBUP_StateHandleCase;
END_VAR
END_METHOD

METHOD CHECKTRANSITION
VAR_INPUT
	ITFSTATESERVER : L_UBUP_IStateServer;
END_VAR
END_METHOD

METHOD FINALIZECYCLE
END_METHOD

METHOD PREPARECYCLE
END_METHOD

METHOD PREPARESTATECHANGE
END_METHOD

METHOD SETADDMODULEINFO
VAR_INPUT
	ESUBCOMPTYPE : UDINT;
	SLICINFO : STRING(10);
END_VAR
END_METHOD

METHOD STIMULATETRANSITION
VAR_INPUT
	ECASE : L_UBUP_StateHandleCase;
END_VAR
END_METHOD

METHOD ALLOCPOINTADR
VAR_OUTPUT
	IERRORID : INT;
END_VAR
END_METHOD

METHOD HANDLEREJECTEDREQUEST : BOOL
VAR_INPUT
	ITFREQUESTANNOUNCED : L_UBUP_IRequest;
END_VAR
VAR_OUTPUT
	ITFALTERNATIVEREQUEST : L_UBUP_IRequest;
END_VAR
END_METHOD

METHOD STATE_01_MOVEABS
VAR_INPUT
	ECASE : L_UBUP_StateHandleCase;
	ISTATESERVER : L_UBUP_IStateServer;
END_VAR
END_METHOD

METHOD STATE_02_MOVEABSCONT
VAR_INPUT
	ECASE : L_UBUP_StateHandleCase;
	ISTATESERVER : L_UBUP_IStateServer;
END_VAR
END_METHOD

METHOD STATE_03_MOVEREL
VAR_INPUT
	ECASE : L_UBUP_StateHandleCase;
	ISTATESERVER : L_UBUP_IStateServer;
END_VAR
END_METHOD

METHOD STATE_04_MOVERELCONT
VAR_INPUT
	ECASE : L_UBUP_StateHandleCase;
	ISTATESERVER : L_UBUP_IStateServer;
END_VAR
END_METHOD

METHOD STATE_05_MOVEVEL
VAR_INPUT
	ECASE : L_UBUP_StateHandleCase;
	ISTATESERVER : L_UBUP_IStateServer;
END_VAR
END_METHOD

METHOD PROFILEGENERATOR
VAR_INPUT
	ITFTECHMODULE : L_TF2P_ITablePositioningBase;
	XEXECUTE : BOOL;
	XCONTINUOUSUPDATE : BOOL;
	LRPOSITION : LREAL;
	LRVELOCITY : LREAL;
	LRENDVELOCITY : LREAL;
	LRACCELERATION : LREAL;
	LRDECELERATION : LREAL;
	LRJERK : LREAL;
	XPOSMODE : BOOL;
	EDIRECTION : MC_DIRECTION;
	EFUNCTIONTYP : L_MC1P_TypeFunction;
END_VAR
VAR_OUTPUT
	XDONE : BOOL;
	XBUSY : BOOL;
	XACTIVE : BOOL;
	XCOMMANDABORTED : BOOL;
	XERROR : BOOL;
	EERRORID : L_IE1P_Error;
END_VAR
VAR_IN_OUT
	AXIS : AXIS_REF;
END_VAR
END_METHOD

METHOD CALC_TP_INTEGRATORSTARTVALUE
END_METHOD

METHOD CALL_STATEENTRYALL
END_METHOD

METHOD CALL_STATEEXITALL
END_METHOD

METHOD CALL_STATEPOSTALL
END_METHOD

METHOD CALL_ALLOCPOINTADR
END_METHOD

METHOD CALL_EXIT_CALLFBS
END_METHOD

METHOD CALL_INIT_CALLFBS
END_METHOD

METHOD CALL_INTERNALCTRL
END_METHOD

METHOD CALL_RESETOUTPUT
END_METHOD

METHOD MAPTMSTATE
VAR_INPUT
	ETMSTATEINTERNAL : L_TB2P_States;
END_VAR
VAR_OUTPUT
	ETMSTATEEXTERNAL : L_TB2P_States;
END_VAR
END_METHOD

(* ---- L_TF2P_TM_VIRTUALMASTERBASE.fb ---- *)
FUNCTION_BLOCK L_TF2P_TM_VIRTUALMASTERBASE EXTENDS L_TB2P_SyncMotionControl
VAR
	TM_VIRTUALMASTERBASECONFIG : L_TB2P_ModuleHandlerConfig;
	PSCINPUT : POINTER TO L_TF2P_VirtualMasterBaseIn;
	PSCOUTPUT : POINTER TO L_TF2P_VirtualMasterBaseOut;
	PPAR : POINTER TO L_TF2P_scPar_TM_VirtualMasterBase;
	PSF : POINTER TO L_TF2P_scSF_TM_VirtualMasterBase;
	PAP : POINTER TO L_TF2P_scAP_TM_VirtualMasterBase;
	SCPAR_INT : L_TF2P_scPar_TM_VirtualMasterBase;
	XACCDECSYNC_INT : BOOL;
	XINTARGETPOS_INT : BOOL;
	LRSTARTPOS_INT : LREAL;
	LRTARGETPOS_INT : LREAL;
	LRSETVEL_LOCK : LREAL;
	EDIRECTION_LOCK : MC_DIRECTION;
	LRMASTERSTARTDISTANCE_INT : LREAL;
	LRMASTERSYNCPOSITION_INT : LREAL;
	LRSLAVESYNCPOSITION_INT : LREAL;
	XVIRTUALMASTERMOVEVELEXECUTE_INT : BOOL;
	XVIRTUALMASTERMOVEABSEXECUTE_INT : BOOL;
	EDIRECTIONCYCLICMOTION : MC_DIRECTION;
	XVIRTUALMASTERMOVERELEXECUTE_INT : BOOL;
	XVIRTUALMASTERHALT_INT : BOOL;
	XVIRTUALMASTERHALT_OLD : BOOL;
	XVIRTUALMASTERHALT_NEXCYCLE : BOOL;
	XVIRTUALMASTERABORT_INT : BOOL;
	XVIRTUALMASTERABORT_OLD : BOOL;
	XVIRTUALMASTERABORT_NEXCYCLE : BOOL;
	XCYCLICMOTIONBUSY_INT : BOOL;
	XCYCLICMOTIONDONE_INT : BOOL;
	XCONTINUOUSMOTIONBUSY_INT : BOOL;
	XCONTINUOUSACTIVE_INT : BOOL;
	XCYCLICACTIVE_INT : BOOL;
	XMOVETOTARGETPOSBUSY_INT : BOOL;
	XMOVETOTARGETPOSDONE_INT : BOOL;
	LRMOVETOTARGETPOS_DIST_INT : LREAL;
	LRCONTINUOUSVEL_INT : LREAL;
	XNOTCONTINUOUS_INT : BOOL;
	WOLDSTATE : WORD;
	XSYNCIN_OLD : BOOL;
	XCONTINUOUS_OLD : BOOL;
	XCYCLE_OLD : BOOL;
	XSTOP_OLD : BOOL;
	XLOADSTARTPOS_OLD : BOOL;
	XOLDENABLE : BOOL;
	XSTARTPOSOUTRANGE : BOOL;
	LRTARGETPOS_SAVE : LREAL;
	XSP_EXECUTE : BOOL;
	XMOVETOTARGETPOSACTIVE : BOOL;
	BYSTEPPERMOVETOTARGETPOS : BYTE;
	LRCYCLELENGTH : LREAL;
	XINVALIDSYNCSLAVEDIRECTION : BOOL;
	XINTERNALCONTR_R_EDGE : R_TRIG;
	FB_SETPOSITION : MC_SetPosition;
	XWARNING_SYNCMODEVELACCREQUIRED : BOOL;
	XWARNING_INVALIDSYNCSLAVEDIRECTION : BOOL;
	XWARNING_MODULOAXISISREQUIRED : BOOL;
	XWARNINGNOVALIDVELOCITYMOVETOTARGETPOS : BOOL;
	FB_CLUTCHEXTENDEDBASE : L_TB2P_ClutchExtendedBase;
	FB_CONTROLSETVALUES : L_MC1P_ControlSetValues;
	XQSPAPPLICATION_OLD : BOOL;
	XSYNCOUTATTARGETPOS : BOOL;
	XSYNCOUTATTARGETPOSACTIVE : BOOL;
	BYSTEPPESYNCOUTATTARGETPOS : BYTE := 0;
	XHALT_OLDER : BOOL;
	XABORT_OLDER : BOOL;
	XWARNINGINVALIDMASTERDIRECTIONINT : BOOL;
	XWARNINGDIRECTIONDISABLEDSYNCINT : BOOL;
	XWARNINGDIRECTIONDISABLEDCONTMOTION : BOOL;
	XWARNINGDIRECTIONDISABLEDCYCLIC : BOOL;
	XWARNINGDIRECTIONDISABLEDCONTMOTION_LOCK : BOOL;
	XWARNINGDIRECTIONDISABLEDCYCLIC_LOCK : BOOL;
END_VAR
END_FUNCTION_BLOCK

METHOD CALL_ALLOCPOINTADR
END_METHOD

METHOD CALL_ERRORHANDLER
END_METHOD

METHOD CALL_FBMETHODS
END_METHOD

METHOD CALL_FB_CLUTCHEXTENDEDBASE
END_METHOD

METHOD CALL_FB_CONTROLSETVALUES
END_METHOD

METHOD CALL_INITROUTINE
END_METHOD

METHOD CALL_INTERNALCTRL
END_METHOD

METHOD CALL_INTERNALCTRLSTATE
END_METHOD

METHOD CALL_MC_SETPOSITION
END_METHOD

METHOD CALL_OUTPUT
END_METHOD

METHOD CALL_REQUESTS_EXT
END_METHOD

METHOD CALL_RESETABCMOVEEXECUTE
END_METHOD

METHOD CALL_RESETCOMMANDS
END_METHOD

METHOD CALL_RESETEXTERNALSTATEABC : BOOL
VAR_INPUT
	FUNSTATE : L_MC1P_ABC_State;
END_VAR
END_METHOD

METHOD CALL_RESETOUTPUT
END_METHOD

METHOD CALL_SETABCMOVEPAR
END_METHOD

METHOD CALL_SETABCMOVESETVEL
END_METHOD

METHOD CALL_SETCLUTCHPOSPAR
END_METHOD

METHOD CALL_SYNCDRIVE
END_METHOD

METHOD SWITCHTOEXTMASTER
END_METHOD

METHOD CALL_ABC_INPUT
END_METHOD

METHOD CALL_ABC_INPUT_PROFILEPARAMETER
END_METHOD

METHOD CALL_CLUTCHOUT
END_METHOD

METHOD CALL_S000_CYCLIC
END_METHOD

METHOD CALL_S002_STANDBY
END_METHOD

METHOD CALL_S030_SYNCHRONISING_POS
END_METHOD

METHOD CALL_S031_POS_IS_SYNCHRONISED
END_METHOD

METHOD CALL_S035_MOVE_TO_TARGET_POS
END_METHOD

METHOD CALL_S060_CONTMOTION
END_METHOD

METHOD CALL_S130_CYCLICMOTION
END_METHOD

METHOD CALL_S996_STOP
END_METHOD

METHOD CALL_S999_ERROR
END_METHOD

METHOD CALL_STATEMACHINE
END_METHOD

METHOD CALL_T000_ALLSTATES
END_METHOD

METHOD CALL_T035_MOVE_TO_TARGET_POS
END_METHOD

METHOD CALL_T060_CONTMOTION
END_METHOD

METHOD CALL_S000_CYCLIC_OUT
END_METHOD

METHOD CALL_S030_SYNCHRONISING_POS_OUT
END_METHOD

METHOD CALL_S031_POS_IS_SYNCHRONISED_OUT
END_METHOD

METHOD CALL_S035_MOVE_TO_TARGET_POS_OUT
END_METHOD

METHOD CALL_S060_CONTMOTION_OUT
END_METHOD

METHOD CALL_S130_CYCLICMOTION_OUT
END_METHOD

METHOD CALL_S999_ERROR_OUT
END_METHOD

METHOD CALL_STATEMACHINE_OUT
END_METHOD

METHOD CALL_T035_MOVE_TO_TARGET_POS_OUT
END_METHOD

(* ---- L_TF2P_VIRTUALMASTER_INTERNAL.fb ---- *)
FUNCTION_BLOCK L_TF2P_VIRTUALMASTER_INTERNAL EXTENDS L_TB2P_TechModuleBase
VAR_INPUT
	XENABLE : BOOL;
	XRESETERROR : BOOL;
	XHALT : BOOL;
	XJOGPOS : BOOL;
	XJOGNEG : BOOL;
	SCPAR : L_TF2P_scPar_VirtualMaster_internal;
	MASTERVALUES : L_MC1P_IAXIS_REF_MASTERVALUES;
	XCONTINUOUS : BOOL;
	XCYCLEEXECUTE : BOOL;
	XLOADSTARTPOS : BOOL;
	LRSETVEL : LREAL := 100;
	XSYNCIN : BOOL;
END_VAR
VAR_OUTPUT
	XENABLED : BOOL;
	ESTATE : L_TB2P_States := L_TB2P_States.DISABLED;
	XERROR : BOOL;
	XWARNING : BOOL;
	EERRORID : L_IE1P_Error;
	VIRTUALMASTERAXIS : L_MC1P_IAXIS_REF_MASTERVALUES;
	LRSETPOSOUT : LREAL;
	LRSETVELOUT : LREAL;
	LRSETACCOUT : LREAL;
	XHALTBUSY : BOOL;
	XHALTDONE : BOOL;
	XJOGGINGBUSY : BOOL;
	XCONTINUOUSMOTIONBUSY : BOOL;
	XCYCLICMOTIONBUSY : BOOL;
	XCYCLICMOTIONDONE : BOOL;
	XMOVETOTARGETPOSBUSY : BOOL;
	XMOVETOTARGETPOSDONE : BOOL;
	XINTARGET : BOOL;
	XACCDECSYNC : BOOL;
	XSYNCHRONISED : BOOL;
END_VAR
VAR_IN_OUT
	AXIS : AXIS_REF;
END_VAR
VAR
	_SCINPUT : L_TF2P_VirtualMasterBaseIn_internal;
	_SCOUTPUT : L_TF2P_VirtualMasterBaseOut_internal;
	_SCINPUTVISU : L_TF2P_VirtualMasterBaseIn_internal;
	_PSCINPUTVISU : POINTER TO L_TF2P_VirtualMasterBaseIn_internal := ADR(_scInputVisu);
	_PSCOUTPUTVISU : POINTER TO L_TF2P_VirtualMasterBaseOut_internal := ADR(_scOutput);
	_PSCPARVISU : POINTER TO L_TF2P_scPar_VirtualMaster_internal := ADR(scPar_int);
	UDIAPPCREDIT : UDINT := 25;
	FB_CLUTCHEXTENDEDBASE : L_TB2P_ClutchExtendedBase;
	FB_FOLLOWSETVALUES : L_MC1P_FollowSetValues;
	MC_POWER : MC_Power;
	MASTERVALUES_INT : L_MC1P_IAXIS_REF_MASTERVALUES;
	FB_L_MC1P_SETAXISREFMASTERVALUES : L_MC1P_SetAxisRefMasterValues;
	READACTUALERRORCODE : L_IE1P_ReadActualErrorCode;
	FBBASE : L_MC1P_Template_ForAxis;
	FBMB : L_MC1P_MoveBasic := STRUCT(wCalcProfileMode := 1);
	EFUNCTIONTYP : L_MC1P_TypeFunction;
	XINTERNALCONTROL_OLD : BOOL;
	SCPAR_INT : L_TF2P_scPar_VirtualMaster_internal;
	LRSTARTPOS_INT : LREAL;
	LRTARGETPOS_INT : LREAL;
	EFBSTATE_INT : L_TB2P_States := L_TB2P_States.DISABLED;
	XSTARTCONTINUOUS_INT : BOOL;
	XSTARTCYCLEEXECUTE_INT : BOOL;
	XSTARTJOGPOS_INT : BOOL;
	XSTARTJOGNEG_INT : BOOL;
	XSTARTHALT_INT : BOOL;
	XENABLEOLD : BOOL;
	XCONTINUOUSOLD : BOOL;
	XCYCLEEXECUTEOLD : BOOL;
	XJOGPOSOLD : BOOL;
	XJOGNEGOLD : BOOL;
	XSYNCINOLD : BOOL;
	XHALTOLD : BOOL;
	XMOVETOTARGETPOSBUSYOLD : BOOL;
	XFBERROR_INT : BOOL;
	XFBERROR_OLD : BOOL;
	XFBWARNING_INT : BOOL;
	EFBERRORID_INT : L_IE1P_Error := 0;
	XCLUTCHACTIVE : BOOL := FALSE;
	XLOADSTARTPOSOLD : BOOL;
	XJOGGINGFLAGPOS : BOOL;
	XJOGGINGFLAGNEG : BOOL;
	XSYNCFLAG : BOOL;
	XCYCLEFLAG : BOOL;
	XCONTINUOUSFLAG : BOOL;
	XHALTFLAG : BOOL;
	XCYCLICDONEFLAG : BOOL;
	XMASTERITFVALID : BOOL;
	BYMASTERID : POINTER TO BYTE;
	XMASTERITFVALID_LOCK : BOOL;
	BYMASTERID_LOCK : POINTER TO BYTE;
	EMASTERTRAVERSINGRANGE : L_MC1P_TraversingRange;
	LRMASTERCYCLELENGTH : LREAL;
	LRSETVELOLD_INT : LREAL;
	PPAR : POINTER TO L_TF2P_scPar_VirtualMaster_internal := ADR(scPar_int);
	XEXECUTEPROFILE_INT : BOOL;
	LRVELOCITY : LREAL;
	LRPOSITION : LREAL;
	LRENDVELOCITY : LREAL;
	LRACC : LREAL;
	LRDEC : LREAL;
	LRJERK : LREAL;
	XPOSMODE : BOOL;
	DIRECTION : MC_DIRECTION := MC_DIRECTION.mcPositiveDirection;
	DONE : BOOL;
	BUSY : BOOL;
	ACTIVE : BOOL;
	COMMANDABORTED : BOOL;
	ERROR : BOOL;
	ERRORID : L_IE1P_Error;
	L_IE1P_SETERROR1 : L_IE1P_SetError;
	XERRORPOSOUTOFCYCLELENGTH : BOOL;
	XERRORPOSOUTOFCYCLELENGTH_OLD : BOOL;
	XJOGRAMPDOWN : BOOL := FALSE;
	XACCDECFLAG : BOOL := FALSE;
	XSTARTNEWCYCLE : BOOL := FALSE;
	TRAVERSINGRANGEOLD : L_MC1P_TraversingRange;
	ESTATEOLD : L_TB2P_States := L_TB2P_States.DISABLED;
	XAXISREADYFORMOTIONOLD : BOOL;
	XDISABLEOLDHALT : BOOL;
	XINTARGETSAVE : BOOL;
	XSTARTMOVETOTARGETPOS : BOOL;
	XMOVETOTARGETPOSZEROVEL : BOOL;
	L_MC1P_GETDIRECTION : L_MC1P_GetDirection;
	_XREADYFORSYNCMOTION : BOOL;
	DWLIMITERCONTROL : DWORD;
END_VAR
END_FUNCTION_BLOCK

METHOD CALL_ALLOCPOINTADR
END_METHOD

METHOD CALL_ERRORHANDLER
END_METHOD

METHOD CALL_ERRORRESETACTIVE
END_METHOD

METHOD CALL_ERRORHANDLER_SCERRORINFO
END_METHOD

METHOD CALL_FB_CLUTCHEXTENDEDBASE
END_METHOD

METHOD CALL_INTERNALCTRL
END_METHOD

METHOD CALL_MASTERVALUESREF
VAR_INPUT
	MASTERVALUES : L_MC1P_IAXIS_REF_MASTERVALUES;
END_VAR
END_METHOD

METHOD CALL_RESETFLAGS
END_METHOD

METHOD CALL_RESETINTERNALCONTROL
END_METHOD

METHOD CALL_RESETOUTPUTS
END_METHOD

METHOD CALL_SETERROR
END_METHOD

METHOD CALL_STATEMACHINE
VAR_IN_OUT
	AXIS : AXIS_REF;
END_VAR
END_METHOD

METHOD CALL_STATEMACHINE_OUT
VAR_IN_OUT
	AXIS : AXIS_REF;
END_VAR
END_METHOD

METHOD GET_PAP : POINTER TO L_TB2P_scAP_TM_MotionControl
END_METHOD

METHOD GET_PPAR : POINTER TO L_TB2P.L_TB2P_scPar_TM_MotionControl
END_METHOD

METHOD GET_PSF : POINTER TO L_TB2P_scSF_TM_MotionControl
END_METHOD

METHOD CALLFUNCTION
END_METHOD

METHOD COPYINPUTS : BOOL
END_METHOD

METHOD COPYOUTPUTS : BOOL
END_METHOD

METHOD FUNCTIONWASCALLEDTWICE : BOOL
VAR_INPUT
	IDX : WORD;
END_VAR
END_METHOD

METHOD HANDLESTANDARDCALL : BOOL
END_METHOD

METHOD SYNCOUTPUTS
VAR_INPUT
	UICOPYOUTPUTFROMIDX : UINT;
	UICOPYOUTPUTTOIDX : UINT;
END_VAR
END_METHOD

(* ---- L_TF2P_VIRTUALMASTERBASE.fb ---- *)
FUNCTION_BLOCK L_TF2P_VIRTUALMASTERBASE EXTENDS L_TB2P_TechModuleBase
VAR_INPUT
	XENABLE : BOOL;
	XENABLEOPERATION : BOOL;
	XRESETERROR : BOOL;
	XQSPAPPLICATION : BOOL;
	XABORT : BOOL;
	XJOGPOS : BOOL;
	XJOGNEG : BOOL;
	XHOMEEXECUTE : BOOL;
	LROVERRIDE : LREAL := 1;
	SCCTRLBASICMOTION : L_TB2P_scCtrlBasicMotion;
	SCPAR : L_TF2P_scPar_VirtualMasterBase;
	SCACCESSPOINTS : L_TF2P_scAP_VirtualMasterBase;
	MASTERVALUES : L_MC1P_IAXIS_REF_MASTERVALUES;
	XCONTINUOUS : BOOL;
	XCYCLEEXECUTE : BOOL;
	XLOADSTARTPOS : BOOL;
	LRSETVEL : LREAL := 10;
	XSYNCIN : BOOL;
END_VAR
VAR_OUTPUT
	XREADYFOROPERATION : BOOL;
	XOPERATIONENABLED : BOOL;
	XREADYFORMOTION : BOOL;
	XERROR : BOOL;
	XWARNING : BOOL;
	EERRORID : L_IE1P_Error;
	XSTOACTIVE : BOOL;
	XQSPACTIVE : BOOL;
	XABORTBUSY : BOOL;
	XABORTDONE : BOOL;
	XJOGGINGBUSY : BOOL;
	XHOMINGBUSY : BOOL;
	XHOMINGDONE : BOOL;
	XISHOMED : BOOL;
	ETMSTATE : L_TB2P_States := L_TB2P_States.DISABLED;
	SCSTATUSBASICMOTION : L_TB2P_scStatusBasicMotion;
	LRACTVEL : LREAL;
	LRSETVELOUT : LREAL;
	LRACTPOS : LREAL;
	LRSETPOSOUT : LREAL;
	LRACTFOLLOWINGERROR : LREAL;
	SCSIGNALFLOW : L_TF2P_scSF_VirtualMasterBase;
	XCONTINUOUSMOTIONBUSY : BOOL;
	XCYCLICMOTIONBUSY : BOOL;
	XCYCLICMOTIONDONE : BOOL;
	XMOVETOTARGETPOSBUSY : BOOL;
	XMOVETOTARGETPOSDONE : BOOL;
	XINTARGET : BOOL;
	XACCDECSYNC : BOOL;
	XSYNCHRONISED : BOOL;
END_VAR
VAR_IN_OUT
	AXIS : AXIS_REF;
END_VAR
VAR
	TM_INT : L_TF2P_TM_VirtualMasterBase := STRUCT(ModuleHandler := ModuleHandler);
	PPAR : POINTER TO L_TF2P_scPar_VirtualMasterBase;
	PPAR_INT : POINTER TO L_TF2P_scPar_VirtualMasterBase;
	_UICALLMFUNIDXINPUT : UINT := 1;
	_UICALLMFUNIDXOUTPUT : UINT := 1;
	_ASCINPUT : ARRAY [1.._MCCall.c_BufferDepthInput] OF L_TF2P_VirtualMasterBaseIn;
	_ASCOUTPUT : ARRAY [1.._MCCall.c_BufferDepthOutput] OF L_TF2P_VirtualMasterBaseOut;
	_ASCPARCORE : ARRAY [1.._MCCall.c_BufferDepthInput] OF L_TF2P_scPar_VirtualMasterBase;
	_ASCACCESSPOINTSCORE : ARRAY [1.._MCCall.c_BufferDepthInput] OF L_TF2P_scAP_VirtualMasterBase;
	_ASCSIGNALFLOWCORE : ARRAY [1.._MCCall.c_BufferDepthOutput] OF L_TF2P_scSF_VirtualMasterBase;
	_MCCALL : L_UM1P_MCCall;
	SCPAR_INT : L_TF2P_scPar_VirtualMasterBase;
	_SCINPUTVISU : L_TF2P_VirtualMasterBaseIn;
	_PSCINPUTVISU : POINTER TO L_TF2P_VirtualMasterBaseIn := ADR(_scInputVisu);
	_PSCOUTPUTVISU : POINTER TO L_TF2P_VirtualMasterBaseOut := ADR(_ascOutput[1]);
	_PSCPARVISU : POINTER TO L_TF2P_scPar_VirtualMasterBase := ADR(scPar_int);
	ITFITECHMODULEINTERNAL : L_TB2P_ITechModuleInternal;
	LRJERKDEC : LREAL;
	LRJOGGINGJERKDEC : LREAL;
	REMAININGTIMEOFPROFILE : LREAL;
	REMAININGTIMEOFPROFILEAVAILABLE : BOOL;
END_VAR
END_FUNCTION_BLOCK

METHOD GET_PAP : POINTER TO L_TB2P_scAP_TM_MotionControl
END_METHOD

METHOD GET_PPAR : POINTER TO L_TB2P.L_TB2P_scPar_TM_MotionControl
END_METHOD

METHOD GET_PSF : POINTER TO L_TB2P_scSF_TM_MotionControl
END_METHOD

METHOD CALLFUNCTION
VAR_INPUT
	UIINPUTDATAIDX : UINT;
	UIOUTPUTDATAIDX : UINT;
END_VAR
END_METHOD

METHOD COPYINPUTS : BOOL
VAR_INPUT
	IDX : WORD;
END_VAR
END_METHOD

METHOD COPYOUTPUTS : BOOL
VAR_INPUT
	IDX : WORD;
END_VAR
END_METHOD

METHOD FUNCTIONWASCALLEDTWICE : BOOL
VAR_INPUT
	IDX : WORD;
END_VAR
END_METHOD

METHOD HANDLESTANDARDCALL : BOOL
END_METHOD

METHOD SYNCOUTPUTS
VAR_INPUT
	UICOPYOUTPUTFROMIDX : UINT;
	UICOPYOUTPUTTOIDX : UINT;
END_VAR
END_METHOD

METHOD CALL_INTERNALCTRL
END_METHOD
